(*
SPDX-FileCopyrightText: c 2026 Oleksandr Tiutyk <trofimich@gmail.com>
SPDX-License-Identifier: MIT
License: https://opensource.org/license/mit
*)

(*!
<summary>Checks the concrete assignment failures and recovery with a matching buffer.</summary>
<description>
Uses one task and stays at a stable address while assertions are bound to this instance.
</description>
*)

{attribute 'no_assign'}
{attribute 'no_explicit_call' := 'do not call this function block directly'}
FUNCTION_BLOCK WideStringBuilderAssignmentFailureTest EXTENDS TOF_Testing.SingleCycleTest
VAR_STAT
	{attribute 'hide'}
	_ClassName : STRING := __POUNAME();
END_VAR
VAR
	_Builder : TOF_Core.WideStringBuilder;
END_VAR

(*!
<summary>Checks the concrete assignment failures and recovery with a matching buffer.</summary>
<description>
The builder is persistent so teardown can release its buffer after an unexpected hook exception.
</description>
*)
METHOD PROTECTED ExecuteTest
VAR
	byteTarget : STRING := 'byte sentinel';
	shortTarget : WSTRING(10) := "keep";
	exactTarget : WSTRING(16);

	exceptionCode : __SYSTEM.ExceptionCode;
	caught : TOF_Core.IException;
	typeException : TOF_Core.IArgumentTypeClassNotSupportedException;
	capacityException : TOF_Core.ITargetVariableMemoryOverflowException;
	copied : BOOL;
END_VAR
_Builder.AppendString255(value := "String1234567890");

// Invoke a wrong-width target and check that the argument is rejected before modification.
__TRY
	_Builder.AssignToString(targetString := byteTarget);
__CATCH(exceptionCode)
	caught := TOF_Core.ExceptionManager.GetLastException(
		exceptionCode := exceptionCode,
		catchPointNamespaceName := NamespaceName,
		catchPointPOUName := __POUNAME(),
		catchPointPosition := __POSITION()
	);
__ENDTRY

Assert.ThatBool(
	actual := __QUERYINTERFACE(caught, typeException),
	message := "AssignToString must report an incompatible STRING target"
).IsTrue();
Assert.ThatBool(
	actual := byteTarget = 'byte sentinel',
	message := "Wrong-width assignment must preserve the target"
).IsTrue();

caught := 0;

// Invoke an undersized WSTRING target and capture the documented capacity exception.
__TRY
	_Builder.AssignToString(targetString := shortTarget);
__CATCH(exceptionCode)
	caught := TOF_Core.ExceptionManager.GetLastException(
		exceptionCode := exceptionCode,
		catchPointNamespaceName := NamespaceName,
		catchPointPOUName := __POUNAME(),
		catchPointPosition := __POSITION()
	);
__ENDTRY

Assert.ThatBool(
	actual := __QUERYINTERFACE(caught, capacityException),
	message := "AssignToString must report insufficient capacity"
).IsTrue();
Assert.ThatBool(
	actual := shortTarget = "keep",
	message := "Capacity rejection must preserve the target"
).IsTrue();

copied := _Builder.AssignToString(targetString := exactTarget);
Assert.ThatBool(
	actual := copied AND_THEN exactTarget = "String1234567890",
	message := "The same builder must still copy successfully into the exact-fit target"
).IsTrue();
END_METHOD

(*!
<summary>Releases the builder buffer before reporting the case result.</summary>
<description>
Safe after partial initialization and after explicit cleanup in the scenario.
</description>
*)
METHOD PROTECTED AfterTest
_Builder.Clear(releaseMemory := TRUE);
END_METHOD

//! <summary>Borrows the concrete class name. Callers must not modify it.</summary>
{attribute 'monitoring' := 'call'}
PROPERTY ClassName : REFERENCE TO STRING
GET
ClassName REF= _ClassName;
END_GET
END_PROPERTY

//! <summary>Borrows the compiler-initialized namespace name. Callers must not modify it.</summary>
{attribute 'monitoring' := 'call'}
PROPERTY NamespaceName : REFERENCE TO STRING
GET
NamespaceName REF= CurrentNamespace.Name;
END_GET
END_PROPERTY

//! <summary>Reports the concrete instance size in bytes.</summary>
{attribute 'monitoring' := 'call'}
PROPERTY SelfSize : ULINT
GET
SelfSize := XSIZEOF(THIS^);
END_GET
END_PROPERTY

END_FUNCTION_BLOCK

(* stored: Version 1.1.0.1
   POU WideStringBuilderAssignmentFailureTest: Id {7b87318e-996d-4822-b9d4-aebcec5cf63c}, SpecialFunc None
   Method ExecuteTest: Id {6640a95c-0973-45a8-91a0-6f19ed6e8409}
   Method AfterTest: Id {e7742bcf-ec5e-4c92-afaf-6990aba9e40a}
   Property ClassName: Id {18d28ce0-6701-488a-b9ba-92c34f37f429}
   Get Get: Id {d97d895a-3ac5-4069-ba89-1406fcd27cf7}
   Property NamespaceName: Id {c6cabf7c-d924-4be6-b2b4-78da98b04585}
   Get Get: Id {557981e1-398f-490c-9aa1-33684f5270e9}
   Property SelfSize: Id {540ca1ef-93dd-49e7-8cb9-46c68e143d22}
   Get Get: Id {935b831a-f36f-4afd-949b-12db2474f576} *)
